      FC_W[1,9] := 0.25226828;
      FC_W[1,10] := -0.62714863;
      FC_W[1,11] := 0.07386149;
      FC_W[1,12] := -0.54759747;
      FC_W[1,13] := 0.00231634;
      FC_W[1,14] := -0.22999668;
      FC_W[1,15] := -0.03627737;
      FC_W[1,16] := -0.00447914;
      FC_W[1,17] := 0.00040707;
      FC_W[1,18] := 0.21295871;
      FC_W[1,19] := 0.21917404;
      FC_W[1,20] := -2.03310800;
      FC_W[1,21] := -0.23101221;
      FC_W[1,22] := 0.59129870;
      FC_W[1,23] := -0.14532049;
      FC_W[1,24] := 0.97670478;
      FC_W[1,25] := -0.18546271;
      FC_W[1,26] := 0.49225003;
      FC_W[1,27] := 0.23357685;
      FC_W[1,28] := -0.05720856;
      FC_W[1,29] := 0.13206857;
      FC_W[1,30] := 0.13029382;
      FC_W[1,31] := -0.28611091;
      FC_W[2,0] := -0.53158796;
      FC_W[2,1] := 2.18231130;
      FC_W[2,2] := 0.15426333;
      FC_W[2,3] := 0.93412578;
      FC_W[2,4] := 0.32678425;
      FC_W[2,5] := -0.29157385;
      FC_W[2,6] := -0.43484834;
      FC_W[2,7] := -0.40118921;
      FC_W[2,8] := -0.73715484;
      FC_W[2,9] := -1.47014546;
      FC_W[2,10] := 0.58461505;
      FC_W[2,11] := 0.72801095;
      FC_W[2,12] := -1.09524512;
      FC_W[2,13] := 0.17780326;
      FC_W[2,14] := 0.55109036;
      FC_W[2,15] := -0.46990421;
      FC_W[2,16] := -0.06730769;
      FC_W[2,17] := 0.69749105;
      FC_W[2,18] := 0.58266920;
      FC_W[2,19] := 0.02913308;
      FC_W[2,20] := 0.18312474;
      FC_W[2,21] := -0.12723203;
      FC_W[2,22] := 1.53492939;
      FC_W[2,23] := 1.18760669;
      FC_W[2,24] := -0.14219350;
      FC_W[2,25] := 0.37169734;
      FC_W[2,26] := -0.22027686;
      FC_W[2,27] := -0.33084327;
      FC_W[2,28] := -0.73663527;
      FC_W[2,29] := 0.07243921;
      FC_W[2,30] := 0.08782770;
      FC_W[2,31] := -0.84531319;
      FC_W[3,0] := 0.55170184;
      FC_W[3,1] := 2.12451887;
      FC_W[3,2] := -0.03638018;
      FC_W[3,3] := -0.92874491;
      FC_W[3,4] := 0.01098804;
      FC_W[3,5] := -0.12194143;
      FC_W[3,6] := -0.20283610;
      FC_W[3,7] := 0.71050656;
      FC_W[3,8] := -0.54710799;
      FC_W[3,9] := 0.84274971;
      FC_W[3,10] := -0.37954244;
      FC_W[3,11] := -0.17364120;
      FC_W[3,12] := 0.44716811;
      FC_W[3,13] := -0.05414552;
      FC_W[3,14] := -0.30617589;
      FC_W[3,15] := 0.00501720;
      FC_W[3,16] := -0.61364305;
      FC_W[3,17] := -0.40598497;
      FC_W[3,18] := 0.24112742;
      FC_W[3,19] := -0.18145135;
      FC_W[3,20] := 0.72023159;
      FC_W[3,21] := 0.31241485;
      FC_W[3,22] := -0.22940150;
      FC_W[3,23] := 0.32834825;
      FC_W[3,24] := -0.47077408;
      FC_W[3,25] := -0.41148546;
      FC_W[3,26] := 0.16142704;
      FC_W[3,27] := -0.05713443;
      FC_W[3,28] := -0.32514808;
      FC_W[3,29] := 0.26252571;
      FC_W[3,30] := 0.50961155;
      FC_W[3,31] := 0.53038257;
      FC_W[4,0] := -0.41400927;
      FC_W[4,1] := 1.33202946;
      FC_W[4,2] := 0.12711546;
      FC_W[4,3] := -0.08963529;
      FC_W[4,4] := 0.24866593;
      FC_W[4,5] := 0.08165067;
      FC_W[4,6] := 0.50525010;
      FC_W[4,7] := 0.82496148;
      FC_W[4,8] := 0.11588583;
      FC_W[4,9] := -0.21680501;
      FC_W[4,10] := 0.62970287;
      FC_W[4,11] := 0.06018925;
      FC_W[4,12] := 0.68656421;
      FC_W[4,13] := -1.21256888;
      FC_W[4,14] := -1.26492715;
      FC_W[4,15] := -0.70575857;
      FC_W[4,16] := -0.17878854;
      FC_W[4,17] := 0.27561840;
      FC_W[4,18] := -0.38193029;
      FC_W[4,19] := 0.25415263;
      FC_W[4,20] := -0.94903797;
      FC_W[4,21] := -0.59143215;
      FC_W[4,22] := -0.27362382;
      FC_W[4,23] := -0.23873141;
      FC_W[4,24] := -1.53285766;
      FC_W[4,25] := -0.27194324;
      FC_W[4,26] := -0.57270604;
      FC_W[4,27] := -0.31816959;
      FC_W[4,28] := 0.51076263;
      FC_W[4,29] := -0.39650953;
      FC_W[4,30] := -0.06086056;
      FC_W[4,31] := -0.04000641;
      FC_W[5,0] := 0.25593293;
      FC_W[5,1] := -0.71731991;
      FC_W[5,2] := 0.62669879;
      FC_W[5,3] := 1.38078809;
      FC_W[5,4] := -0.12516685;
      FC_W[5,5] := -0.90641493;
      FC_W[5,6] := -0.39019036;
      FC_W[5,7] := -0.45447922;
      FC_W[5,8] := 0.01198741;
      FC_W[5,9] := -0.21863569;
      FC_W[5,10] := 0.71772867;
      FC_W[5,11] := 0.27339056;
      FC_W[5,12] := 0.20110083;
      FC_W[5,13] := -0.13613328;
      FC_W[5,14] := -2.24843359;
      FC_W[5,15] := 0.12153642;
      FC_W[5,16] := 0.93278831;
      FC_W[5,17] := -0.95549434;
      FC_W[5,18] := 0.26438603;
      FC_W[5,19] := 0.19650064;
      FC_W[5,20] := -0.06620517;
      FC_W[5,21] := 0.29557747;
      FC_W[5,22] := 1.31400585;
      FC_W[5,23] := -0.15871854;
      FC_W[5,24] := 0.40522489;
      FC_W[5,25] := 0.03414011;
      FC_W[5,26] := -0.38867807;
      FC_W[5,27] := -0.81741858;
      FC_W[5,28] := 1.06798649;
      FC_W[5,29] := 3.75573659;
      FC_W[5,30] := -0.51656634;
      FC_W[5,31] := -0.28770104;
      FC_W[6,0] := -0.99143010;
      FC_W[6,1] := 0.29992977;
      FC_W[6,2] := 1.43284762;
      FC_W[6,3] := -0.34655777;
      FC_W[6,4] := -0.12928130;
      FC_W[6,5] := 0.15707546;
      FC_W[6,6] := -0.63261580;
      FC_W[6,7] := -0.29724568;
      FC_W[6,8] := 0.13134219;
      FC_W[6,9] := -1.04233253;
      FC_W[6,10] := 0.53604454;
      FC_W[6,11] := -0.18040322;
      FC_W[6,12] := 0.16615772;
      FC_W[6,13] := -0.40025923;
      FC_W[6,14] := -1.54933608;
      FC_W[6,15] := 0.41574958;
      FC_W[6,16] := 0.35386816;
      FC_W[6,17] := -0.45704508;
      FC_W[6,18] := 0.60151654;
      FC_W[6,19] := -0.67978704;
      FC_W[6,20] := 0.15072536;
      FC_W[6,21] := -0.42846721;
      FC_W[6,22] := -0.85208124;
      FC_W[6,23] := -0.05353868;
      FC_W[6,24] := 0.86764193;
      FC_W[6,25] := -0.24695079;
      FC_W[6,26] := 0.82921457;
      FC_W[6,27] := -1.08330154;
      FC_W[6,28] := 0.22054735;
      FC_W[6,29] := -0.23250555;
      FC_W[6,30] := 0.84133679;
      FC_W[6,31] := -0.10032179;
      FC_W[7,0] := 0.30265906;
      FC_W[7,1] := 2.08623362;
      FC_W[7,2] := 0.06350639;
      FC_W[7,3] := -1.09427238;
      FC_W[7,4] := -0.02930364;
      FC_W[7,5] := 0.24324393;
      FC_W[7,6] := 0.16107884;
      FC_W[7,7] := -0.00278581;
      FC_W[7,8] := 0.11302312;
      FC_W[7,9] := 0.10457820;
      FC_W[7,10] := -0.14860652;
      FC_W[7,11] := -0.10135441;
      FC_W[7,12] := 1.27947247;
      FC_W[7,13] := -0.08310315;
      FC_W[7,14] := -0.41487727;
      FC_W[7,15] := 0.17592667;
      FC_W[7,16] := -0.25739285;
      FC_W[7,17] := 0.24304490;
      FC_W[7,18] := -0.47447765;
      FC_W[7,19] := -0.28621474;
      FC_W[7,20] := 0.67906636;
      FC_W[7,21] := -0.40683922;
      FC_W[7,22] := -0.50886548;
      FC_W[7,23] := 0.06748977;
      FC_W[7,24] := -0.28961775;
      FC_W[7,25] := -0.11677405;
      FC_W[7,26] := 0.16660805;
      FC_W[7,27] := 0.34886500;
      FC_W[7,28] := -0.65834177;
      FC_W[7,29] := 0.30940986;
      FC_W[7,30] := -0.04497011;
      FC_W[7,31] := 0.22881326;
      FC_W[8,0] := 0.23515312;
      FC_W[8,1] := 2.35528612;
      FC_W[8,2] := 0.12001805;
      FC_W[8,3] := 0.60647392;
      FC_W[8,4] := -0.31542465;
      FC_W[8,5] := -0.26584071;
      FC_W[8,6] := 0.15293968;
      FC_W[8,7] := 0.19515641;
      FC_W[8,8] := -0.34400198;
      FC_W[8,9] := 0.12394456;
      FC_W[8,10] := 0.06283668;
      FC_W[8,11] := -0.67132694;
      FC_W[8,12] := -1.10496128;
      FC_W[8,13] := -0.33543864;
      FC_W[8,14] := 0.34250832;
      FC_W[8,15] := 0.11089487;
      FC_W[8,16] := 0.27817380;
      FC_W[8,17] := -0.27934778;
      FC_W[8,18] := 1.01753807;
      FC_W[8,19] := -0.14856282;
      FC_W[8,20] := 1.15498221;
      FC_W[8,21] := 0.31782010;
      FC_W[8,22] := -0.57135326;
      FC_W[8,23] := -0.27457404;
      FC_W[8,24] := -0.01912341;
      FC_W[8,25] := 0.07636409;
      FC_W[8,26] := -0.05262562;
      FC_W[8,27] := 0.01281669;
      FC_W[8,28] := 1.45306993;
      FC_W[8,29] := 0.01643326;
      FC_W[8,30] := 0.02226772;
      FC_W[8,31] := 0.16109315;
      FC_W[9,0] := 0.16771235;
      FC_W[9,1] := 2.17360902;
      FC_W[9,2] := 0.13744619;
      FC_W[9,3] := -0.45034087;
      FC_W[9,4] := -0.18103811;
      FC_W[9,5] := 0.19206211;
      FC_W[9,6] := 0.29432642;
      FC_W[9,7] := -0.29548097;
      FC_W[9,8] := 0.26934287;
      FC_W[9,9] := -0.23640421;
      FC_W[9,10] := 0.08889509;
      FC_W[9,11] := -0.29550803;
      FC_W[9,12] := 0.70984375;
      FC_W[9,13] := -0.18878627;
      FC_W[9,14] := -0.16082951;
      FC_W[9,15] := 0.28989646;
      FC_W[9,16] := 0.17481117;
      FC_W[9,17] := 0.31475934;
      FC_W[9,18] := -0.19749227;
      FC_W[9,19] := -0.29642978;
      FC_W[9,20] := 0.85720885;
      FC_W[9,21] := -0.43476731;
      FC_W[9,22] := -0.67719740;
      FC_W[9,23] := -0.20220257;
      FC_W[9,24] := -0.05126322;
      FC_W[9,25] := 0.10412872;
      FC_W[9,26] := 0.06379344;
      FC_W[9,27] := 0.43333077;
      FC_W[9,28] := 0.06093162;
      FC_W[9,29] := 0.21085459;
      FC_W[9,30] := -0.27212784;
      FC_W[9,31] := 0.04487327;
      FC_W[10,0] := 0.55635911;
      FC_W[10,1] := 1.71071684;
      FC_W[10,2] := -0.98758829;
      FC_W[10,3] := -1.20704234;
      FC_W[10,4] := 0.70373571;
      FC_W[10,5] := -0.49822235;
      FC_W[10,6] := -0.34963137;
      FC_W[10,7] := -0.04954350;
      FC_W[10,8] := 0.57998538;
      FC_W[10,9] := -0.12894104;
      FC_W[10,10] := 0.17007013;
      FC_W[10,11] := 0.22826548;
      FC_W[10,12] := 0.52343917;
      FC_W[10,13] := 0.24545214;
      FC_W[10,14] := 0.32942688;
      FC_W[10,15] := 0.31240448;
      FC_W[10,16] := -0.23860073;
      FC_W[10,17] := 0.84877467;
      FC_W[10,18] := -0.03334466;
      FC_W[10,19] := -0.08059564;
      FC_W[10,20] := -0.50759733;
      FC_W[10,21] := 0.57257271;
      FC_W[10,22] := -0.54642487;
      FC_W[10,23] := 0.07352713;
      FC_W[10,24] := 0.81966442;
      FC_W[10,25] := -0.40594006;
      FC_W[10,26] := -0.35969523;
      FC_W[10,27] := 1.14789081;
      FC_W[10,28] := 0.64354020;
      FC_W[10,29] := 1.38284671;
      FC_W[10,30] := -0.42893896;
      FC_W[10,31] := 0.09688565;
      FC_W[11,0] := -0.43645921;
      FC_W[11,1] := 0.23312488;
      FC_W[11,2] := -0.23381421;
      FC_W[11,3] := 1.35307658;
      FC_W[11,4] := 0.06825005;
      FC_W[11,5] := 0.04006363;
      FC_W[11,6] := -0.30487701;
      FC_W[11,7] := -0.04899468;
      FC_W[11,8] := -0.69408715;
      FC_W[11,9] := 0.32083067;
      FC_W[11,10] := -1.27051854;
      FC_W[11,11] := -0.28955328;
      FC_W[11,12] := 0.94128507;
      FC_W[11,13] := -0.04163137;
      FC_W[11,14] := -0.19035473;
      FC_W[11,15] := 1.00236845;
      FC_W[11,16] := 1.06163549;
      FC_W[11,17] := 0.45048153;
      FC_W[11,18] := 0.19175214;
      FC_W[11,19] := -0.00000184;
      FC_W[11,20] := -0.00385919;
      FC_W[11,21] := -0.25575012;
      FC_W[11,22] := 0.63028401;
      FC_W[11,23] := 0.23347531;
      FC_W[11,24] := 0.62187344;
      FC_W[11,25] := -0.06846938;
      FC_W[11,26] := -0.08085597;
      FC_W[11,27] := 0.08367075;
      FC_W[11,28] := 0.07401622;
      FC_W[11,29] := -0.68332726;
      FC_W[11,30] := 0.36182699;
      FC_W[11,31] := 0.09208941;
      FC_W[12,0] := -0.12697175;
      FC_W[12,1] := 0.54007989;
      FC_W[12,2] := -0.23235552;
      FC_W[12,3] := 1.02737308;
      FC_W[12,4] := -0.21164975;
      FC_W[12,5] := -0.18848586;
      FC_W[12,6] := -0.31116375;
      FC_W[12,7] := 0.18885162;
      FC_W[12,8] := 0.26512960;
      FC_W[12,9] := 0.64287508;
      FC_W[12,10] := 0.17899334;
      FC_W[12,11] := 0.11003251;
      FC_W[12,12] := 0.97311103;
      FC_W[12,13] := 0.04088512;
      FC_W[12,14] := 0.28795946;
      FC_W[12,15] := 1.57381439;
      FC_W[12,16] := 0.84596854;
      FC_W[12,17] := -0.53194338;
      FC_W[12,18] := 0.83031321;
      FC_W[12,19] := 0.19111450;
      FC_W[12,20] := -0.29391897;
      FC_W[12,21] := -0.53817254;
      FC_W[12,22] := 1.39124548;
      FC_W[12,23] := 0.21961257;
      FC_W[12,24] := 0.63080877;
      FC_W[12,25] := -0.13176970;
      FC_W[12,26] := 0.19578983;
      FC_W[12,27] := 0.07251017;
      FC_W[12,28] := 0.15489395;
      FC_W[12,29] := -0.56836164;
      FC_W[12,30] := 0.24469846;
      FC_W[12,31] := -0.29308897;
      FC_W[13,0] := 2.20791268;
      FC_W[13,1] := -1.10374355;
      FC_W[13,2] := -0.24162126;
      FC_W[13,3] := 0.77374041;
      FC_W[13,4] := -1.13711357;
      FC_W[13,5] := -1.31870210;
      FC_W[13,6] := 0.47841373;
      FC_W[13,7] := -0.16105147;
      FC_W[13,8] := -0.35249650;
      FC_W[13,9] := -0.42332867;
      FC_W[13,10] := -1.55202627;
      FC_W[13,11] := 1.01507616;
      FC_W[13,12] := -0.63866675;
      FC_W[13,13] := -0.71099406;
      FC_W[13,14] := -0.48592618;
      FC_W[13,15] := -0.37993100;
      FC_W[13,16] := 0.18940821;
      FC_W[13,17] := -0.05538184;
      FC_W[13,18] := -0.14446187;
      FC_W[13,19] := 0.44147074;
      FC_W[13,20] := -0.71370798;
      FC_W[13,21] := -1.35824025;
      FC_W[13,22] := -0.32107875;
      FC_W[13,23] := -0.66948777;
      FC_W[13,24] := 0.46409652;
      FC_W[13,25] := -0.56385392;
      FC_W[13,26] := 1.45479858;
      FC_W[13,27] := 1.22730565;
      FC_W[13,28] := -0.70979494;
      FC_W[13,29] := 0.23732866;
      FC_W[13,30] := 0.40240869;
      FC_W[13,31] := -0.91399556;
      FC_W[14,0] := -0.07104833;
      FC_W[14,1] := -0.28022146;
      FC_W[14,2] := -0.67785078;
      FC_W[14,3] := 0.19481595;
      FC_W[14,4] := -0.03060088;
      FC_W[14,5] := -0.20427652;
      FC_W[14,6] := 0.04726106;
      FC_W[14,7] := 1.98258340;
      FC_W[14,8] := 4.40404320;
      FC_W[14,9] := -1.24794614;
      FC_W[14,10] := -1.24316883;
      FC_W[14,11] := -1.68179226;
      FC_W[14,12] := -0.29661027;
      FC_W[14,13] := 0.01353078;
      FC_W[14,14] := -0.41424713;
      FC_W[14,15] := 0.58704215;
      FC_W[14,16] := -1.78230023;
      FC_W[14,17] := 1.53948402;
      FC_W[14,18] := -0.07893131;
      FC_W[14,19] := -3.22760653;
      FC_W[14,20] := 0.56132263;
      FC_W[14,21] := 0.12644786;
      FC_W[14,22] := 1.26095736;
      FC_W[14,23] := -0.00488345;
      FC_W[14,24] := 0.29457206;
      FC_W[14,25] := -1.28626144;
      FC_W[14,26] := -0.26738542;
      FC_W[14,27] := -0.44110236;
      FC_W[14,28] := -0.43122882;
      FC_W[14,29] := -0.00431219;
      FC_W[14,30] := -0.40952465;
      FC_W[14,31] := -0.30441639;
      FC_W[15,0] := 0.20250924;
      FC_W[15,1] := 0.43626478;
      FC_W[15,2] := 0.27463222;
      FC_W[15,3] := 0.37211508;
      FC_W[15,4] := -0.03340056;
      FC_W[15,5] := -0.06623933;
      FC_W[15,6] := -0.24864028;
      FC_W[15,7] := -0.58677751;
      FC_W[15,8] := -0.61499745;
      FC_W[15,9] := 0.54579276;
      FC_W[15,10] := -0.19726747;
      FC_W[15,11] := 0.12831730;
      FC_W[15,12] := 0.61062902;
      FC_W[15,13] := -0.02127237;
      FC_W[15,14] := 0.21842071;
      FC_W[15,15] := -0.17562330;
      FC_W[15,16] := 0.38656747;
      FC_W[15,17] := 0.59372723;
      FC_W[15,18] := 0.24492693;
      FC_W[15,19] := -1.01225615;
      FC_W[15,20] := -0.01717149;
      FC_W[15,21] := 0.54135400;
      FC_W[15,22] := 1.04819000;
      FC_W[15,23] := -1.09988487;
      FC_W[15,24] := -0.29471993;
      FC_W[15,25] := 0.78609461;
      FC_W[15,26] := 0.23125337;
      FC_W[15,27] := -0.02700599;
      FC_W[15,28] := 0.42768958;
      FC_W[15,29] := -0.29631129;
      FC_W[15,30] := 1.83250082;
      FC_W[15,31] := -0.43059009;
      FC_W[16,0] := -0.37697601;
      FC_W[16,1] := -0.19721903;
      FC_W[16,2] := -0.13793600;
      FC_W[16,3] := 0.07084525;
      FC_W[16,4] := 0.47389659;
      FC_W[16,5] := 0.68528003;
      FC_W[16,6] := 1.65266597;
      FC_W[16,7] := -0.24744993;
      FC_W[16,8] := 1.25457382;
      FC_W[16,9] := 1.49639773;
      FC_W[16,10] := 0.50168604;
      FC_W[16,11] := -0.50251526;
      FC_W[16,12] := -0.00292949;
      FC_W[16,13] := -0.70094889;
      FC_W[16,14] := 0.17360571;
      FC_W[16,15] := -0.58291054;
      FC_W[16,16] := 0.50401050;
      FC_W[16,17] := -1.54409647;
      FC_W[16,18] := -1.89241540;
      FC_W[16,19] := -0.33420387;
      FC_W[16,20] := 0.63442737;
      FC_W[16,21] := -0.10250572;
      FC_W[16,22] := -0.74442780;
      FC_W[16,23] := 2.23745084;
      FC_W[16,24] := 0.97562188;
      FC_W[16,25] := -0.53874046;
      FC_W[16,26] := 0.44360429;
      FC_W[16,27] := 0.48179910;
      FC_W[16,28] := 1.56847930;
      FC_W[16,29] := 0.12322044;
      FC_W[16,30] := 0.58041352;
      FC_W[16,31] := -2.92400813;
      FC_W[17,0] := -0.28855094;
      FC_W[17,1] := -0.73520070;
      FC_W[17,2] := -0.58204508;
      FC_W[17,3] := -2.53923368;
      FC_W[17,4] := 0.04207829;
      FC_W[17,5] := 0.34026721;
      FC_W[17,6] := 0.83833164;
      FC_W[17,7] := 1.37610734;
      FC_W[17,8] := -0.48114690;
      FC_W[17,9] := 0.80318284;
      FC_W[17,10] := 1.40226424;
      FC_W[17,11] := 1.19034028;
      FC_W[17,12] := -1.82810128;
      FC_W[17,13] := 0.07092776;
      FC_W[17,14] := -0.24957196;
      FC_W[17,15] := 0.41651461;
      FC_W[17,16] := 2.31544805;
      FC_W[17,17] := -0.29625085;
      FC_W[17,18] := 0.43194380;
      FC_W[17,19] := -2.91967225;
      FC_W[17,20] := 0.48595843;
      FC_W[17,21] := -0.95144910;
      FC_W[17,22] := -0.56275243;
      FC_W[17,23] := 0.17238346;
      FC_W[17,24] := 0.18526348;
      FC_W[17,25] := -1.61428738;
      FC_W[17,26] := -0.85377961;
      FC_W[17,27] := -0.13946605;
      FC_W[17,28] := -0.68767577;
      FC_W[17,29] := 0.88757920;
      FC_W[17,30] := -1.37992692;
      FC_W[17,31] := -0.30283210;
      FC_W[18,0] := -0.60211664;
      FC_W[18,1] := -0.47432238;
      FC_W[18,2] := 0.49715492;
      FC_W[18,3] := -1.05803704;
      FC_W[18,4] := 0.31516069;
      FC_W[18,5] := 0.60292727;
      FC_W[18,6] := -1.12411284;
      FC_W[18,7] := -0.81225699;
      FC_W[18,8] := 0.22442850;
      FC_W[18,9] := -0.31069636;
      FC_W[18,10] := -0.39883116;
      FC_W[18,11] := -0.00383187;
      FC_W[18,12] := -1.32017577;
      FC_W[18,13] := 0.76117158;
      FC_W[18,14] := -0.59863925;
      FC_W[18,15] := 2.91382790;
      FC_W[18,16] := -0.31635019;
      FC_W[18,17] := -0.69926184;
      FC_W[18,18] := 0.44085792;
      FC_W[18,19] := -0.27446097;
      FC_W[18,20] := 0.68643546;
      FC_W[18,21] := -1.84294975;
      FC_W[18,22] := -0.20962636;
      FC_W[18,23] := -0.22959881;
      FC_W[18,24] := 0.18067747;
      FC_W[18,25] := 0.47698760;
      FC_W[18,26] := -3.78073096;
      FC_W[18,27] := 0.82570255;
      FC_W[18,28] := -0.23815499;
      FC_W[18,29] := 1.09470105;
      FC_W[18,30] := 1.66854107;
      FC_W[18,31] := -0.13462155;
      FC_W[19,0] := 0.44800782;
      FC_W[19,1] := 0.06498748;
      FC_W[19,2] := -0.06952048;
      FC_W[19,3] := -0.51742721;
      FC_W[19,4] := -0.09736256;
      FC_W[19,5] := -0.37422362;
      FC_W[19,6] := -0.15245904;
      FC_W[19,7] := 0.63320434;
      FC_W[19,8] := 1.04222059;
      FC_W[19,9] := 0.06480665;
      FC_W[19,10] := 0.35045585;
      FC_W[19,11] := -0.40922517;
      FC_W[19,12] := -0.08025740;
      FC_W[19,13] := 0.05562712;
      FC_W[19,14] := 0.10890836;
      FC_W[19,15] := -0.13707444;
      FC_W[19,16] := 1.62350214;
      FC_W[19,17] := 0.41023293;
      FC_W[19,18] := 0.34094810;
      FC_W[19,19] := 0.31232962;
      FC_W[19,20] := -0.14682344;
      FC_W[19,21] := 0.48118156;
      FC_W[19,22] := 0.78214991;
      FC_W[19,23] := 0.03551027;
      FC_W[19,24] := -0.44571006;
      FC_W[19,25] := -0.08649512;
      FC_W[19,26] := 0.47158131;
      FC_W[19,27] := -0.36406398;
      FC_W[19,28] := -0.22915788;
      FC_W[19,29] := 0.01263516;
      FC_W[19,30] := 0.57616603;
      FC_W[19,31] := 0.12845607;
      FC_W[20,0] := 0.55101711;
      FC_W[20,1] := 0.35684553;
      FC_W[20,2] := -0.92210096;
      FC_W[20,3] := 0.13750382;
      FC_W[20,4] := 0.01511240;
      FC_W[20,5] := -0.63257527;
      FC_W[20,6] := 1.40384579;
      FC_W[20,7] := -0.21248135;
      FC_W[20,8] := -0.16805060;
      FC_W[20,9] := -0.11867571;
      FC_W[20,10] := -0.39359516;
      FC_W[20,11] := -0.15843204;
      FC_W[20,12] := 0.22070603;
      FC_W[20,13] := 0.71381277;
      FC_W[20,14] := -0.11454471;
      FC_W[20,15] := -0.38763249;
      FC_W[20,16] := -0.09213293;
      FC_W[20,17] := -0.03829917;
      FC_W[20,18] := -0.25112540;
      FC_W[20,19] := 0.09202781;
      FC_W[20,20] := -0.79897386;
      FC_W[20,21] := 0.14058812;
      FC_W[20,22] := -0.30311379;
      FC_W[20,23] := -0.43297794;
      FC_W[20,24] := 0.11171950;
      FC_W[20,25] := 0.17598327;
      FC_W[20,26] := -0.82704544;
      FC_W[20,27] := -0.20293660;
      FC_W[20,28] := -0.50960398;
      FC_W[20,29] := -0.13715295;
      FC_W[20,30] := -0.20570764;
      FC_W[20,31] := -0.22419536;
      FC_W[21,0] := -1.38703454;
      FC_W[21,1] := 0.13443221;
      FC_W[21,2] := 1.65575707;
      FC_W[21,3] := -0.30523026;
      FC_W[21,4] := 0.20814605;
      FC_W[21,5] := 0.44282535;
      FC_W[21,6] := -0.18247518;
      FC_W[21,7] := 0.68251020;
      FC_W[21,8] := -0.51809436;
      FC_W[21,9] := -0.59682101;
      FC_W[21,10] := 0.32860571;
      FC_W[21,11] := -0.65614474;
      FC_W[21,12] := -0.12320014;
      FC_W[21,13] := 1.67703843;
      FC_W[21,14] := 0.01895689;
      FC_W[21,15] := 0.41568109;
      FC_W[21,16] := 0.12311991;
      FC_W[21,17] := -0.85774213;
      FC_W[21,18] := -0.30047303;
      FC_W[21,19] := -0.33377433;
      FC_W[21,20] := 0.02386909;
      FC_W[21,21] := -0.03189978;
      FC_W[21,22] := 0.33781007;
      FC_W[21,23] := -0.20913075;
      FC_W[21,24] := -0.16453424;
      FC_W[21,25] := -0.14679955;
      FC_W[21,26] := 0.59973520;
      FC_W[21,27] := 0.48085397;
      FC_W[21,28] := 0.24753553;
      FC_W[21,29] := -0.01857807;
      FC_W[21,30] := 0.12446254;
      FC_W[21,31] := 0.10629370;
      FC_W[22,0] := 0.19716617;
      FC_W[22,1] := 0.13620606;
      FC_W[22,2] := 0.04876109;
      FC_W[22,3] := 0.23500557;
      FC_W[22,4] := 0.64577067;
      FC_W[22,5] := 0.25040030;
      FC_W[22,6] := 0.29043925;
      FC_W[22,7] := 0.85402560;
      FC_W[22,8] := 0.06459093;
      FC_W[22,9] := -1.23667681;
      FC_W[22,10] := -0.05787567;
      FC_W[22,11] := 0.74056232;
      FC_W[22,12] := 0.22630619;
      FC_W[22,13] := -0.10364483;
      FC_W[22,14] := -0.08892694;
      FC_W[22,15] := -0.34050211;
      FC_W[22,16] := 0.65094274;
      FC_W[22,17] := -1.17275202;
      FC_W[22,18] := -0.78813517;
      FC_W[22,19] := 0.34167442;
      FC_W[22,20] := 0.37342751;
      FC_W[22,21] := 0.12655480;
      FC_W[22,22] := 0.14093940;
      FC_W[22,23] := -0.97658986;
      FC_W[22,24] := 0.29666159;
      FC_W[22,25] := -0.95207864;
      FC_W[22,26] := -0.25645512;
      FC_W[22,27] := 0.21099935;
      FC_W[22,28] := -0.17070027;
      FC_W[22,29] := -0.15547353;
      FC_W[22,30] := 0.05844394;
      FC_W[22,31] := -0.35387653;
      FC_W[23,0] := 2.36117458;
      FC_W[23,1] := -0.27253562;
      FC_W[23,2] := -0.44734445;
      FC_W[23,3] := 0.43230754;
      FC_W[23,4] := 2.77088666;
      FC_W[23,5] := -1.15746760;
      FC_W[23,6] := -0.15780434;
      FC_W[23,7] := -0.08052579;
      FC_W[23,8] := -1.13770092;
      FC_W[23,9] := 0.34222582;
      FC_W[23,10] := -0.76248449;
      FC_W[23,11] := -0.31606591;
      FC_W[23,12] := -0.26905468;
      FC_W[23,13] := -0.65461212;
      FC_W[23,14] := 0.29336941;
      FC_W[23,15] := -0.56090289;
      FC_W[23,16] := -0.30688983;
      FC_W[23,17] := 0.29983157;
      FC_W[23,18] := -0.73118234;
      FC_W[23,19] := -0.10799882;
      FC_W[23,20] := -0.22133076;
      FC_W[23,21] := -1.62908876;
      FC_W[23,22] := 0.32420984;
      FC_W[23,23] := 0.12469828;
      FC_W[23,24] := 0.86695164;
      FC_W[23,25] := 0.00903137;
      FC_W[23,26] := 1.11415207;
      FC_W[23,27] := -0.62709349;
      FC_W[23,28] := -0.02971547;
      FC_W[23,29] := -0.25179407;
      FC_W[23,30] := -0.06880520;
      FC_W[23,31] := 0.58122498;
      FC_W[24,0] := 0.07595386;
      FC_W[24,1] := 0.17389667;
      FC_W[24,2] := -0.13460560;
      FC_W[24,3] := 0.23620439;
      FC_W[24,4] := 0.71178508;
      FC_W[24,5] := 0.42975000;
      FC_W[24,6] := 0.46598688;
      FC_W[24,7] := 1.36021495;
      FC_W[24,8] := 0.10479560;
      FC_W[24,9] := -0.78181171;
      FC_W[24,10] := -0.17630832;
      FC_W[24,11] := 0.88054228;
      FC_W[24,12] := 0.23260193;
      FC_W[24,13] := -0.07906808;
      FC_W[24,14] := 0.03967582;
      FC_W[24,15] := -0.41637811;
      FC_W[24,16] := 0.38345000;
      FC_W[24,17] := -0.55840528;
      FC_W[24,18] := -0.90066504;
      FC_W[24,19] := 0.97068053;
      FC_W[24,20] := 0.60454738;
      FC_W[24,21] := 0.02299176;
      FC_W[24,22] := 0.09866967;
      FC_W[24,23] := -1.46094978;
      FC_W[24,24] := 0.38187879;
      FC_W[24,25] := -1.42997479;
      FC_W[24,26] := -0.37488067;
      FC_W[24,27] := -0.04411485;
      FC_W[24,28] := -0.29138446;
      FC_W[24,29] := -0.07532097;
      FC_W[24,30] := -0.00954079;
      FC_W[24,31] := -0.99948364;
      FC_W[25,0] := 0.08445936;
      FC_W[25,1] := 0.16368021;
      FC_W[25,2] := -0.11429817;
      FC_W[25,3] := 0.25485840;
      FC_W[25,4] := 0.72819227;
      FC_W[25,5] := 0.42307603;
      FC_W[25,6] := 0.45525894;
      FC_W[25,7] := 1.32385421;
      FC_W[25,8] := 0.11924174;
      FC_W[25,9] := -0.79466659;
      FC_W[25,10] := -0.16143492;
      FC_W[25,11] := 0.87378216;
      FC_W[25,12] := 0.22462815;
      FC_W[25,13] := -0.08033443;
      FC_W[25,14] := 0.01655862;
      FC_W[25,15] := -0.40789300;
      FC_W[25,16] := 0.40738490;
      FC_W[25,17] := -0.57628548;
      FC_W[25,18] := -0.88914770;
      FC_W[25,19] := 0.94886303;
      FC_W[25,20] := 0.60112166;
      FC_W[25,21] := 0.02799439;
      FC_W[25,22] := 0.08625803;
      FC_W[25,23] := -1.44966817;
      FC_W[25,24] := 0.37795368;
      FC_W[25,25] := -1.41334343;
      FC_W[25,26] := -0.38357916;
      FC_W[25,27] := -0.01546234;
      FC_W[25,28] := -0.29737470;
      FC_W[25,29] := -0.08744591;
      FC_W[25,30] := -0.01248721;
      FC_W[25,31] := -0.99227226;
      FC_W[26,0] := 2.38675141;
      FC_W[26,1] := 0.10531798;
      FC_W[26,2] := 0.00214429;
      FC_W[26,3] := 0.29302251;
      FC_W[26,4] := -0.95878249;
      FC_W[26,5] := -0.62310410;
      FC_W[26,6] := -0.31759438;
      FC_W[26,7] := 0.11338235;
      FC_W[26,8] := -0.31615138;
      FC_W[26,9] := -1.49054682;
      FC_W[26,10] := 0.93792856;
      FC_W[26,11] := 0.87154341;
      FC_W[26,12] := 0.41643369;
      FC_W[26,13] := -1.12895298;
      FC_W[26,14] := -0.42944503;
      FC_W[26,15] := -0.59216714;
      FC_W[26,16] := 0.45720932;
      FC_W[26,17] := -0.10903971;
      FC_W[26,18] := -1.34624648;
      FC_W[26,19] := -0.30879995;
      FC_W[26,20] := 0.24794732;
      FC_W[26,21] := 0.29367086;
      FC_W[26,22] := 0.73384720;
      FC_W[26,23] := 0.23941633;
      FC_W[26,24] := 0.97845572;
      FC_W[26,25] := -0.83140624;
      FC_W[26,26] := -1.05813015;
      FC_W[26,27] := -0.12844378;
      FC_W[26,28] := 0.53951097;
      FC_W[26,29] := -0.46631601;
      FC_W[26,30] := -0.12978332;
      FC_W[26,31] := 0.57293302;
      FC_W[27,0] := -0.82125789;
      FC_W[27,1] := 0.24535166;
      FC_W[27,2] := 2.14815331;
      FC_W[27,3] := 0.07394390;
      FC_W[27,4] := 0.37535343;
      FC_W[27,5] := 0.20946552;
      FC_W[27,6] := -0.22952469;
      FC_W[27,7] := 0.21198778;
      FC_W[27,8] := 0.45519185;
      FC_W[27,9] := 0.43655413;
      FC_W[27,10] := 0.14163223;
      FC_W[27,11] := 0.37753379;
      FC_W[27,12] := -0.03609978;
      FC_W[27,13] := 1.92808294;
      FC_W[27,14] := 0.01438947;
      FC_W[27,15] := 0.12405793;
      FC_W[27,16] := 0.13592151;
      FC_W[27,17] := 0.25425518;
      FC_W[27,18] := -0.02739565;
      FC_W[27,19] := -0.02477069;
      FC_W[27,20] := 0.06481469;
      FC_W[27,21] := 0.01653567;
      FC_W[27,22] := -0.02758124;
      FC_W[27,23] := 0.17188995;
      FC_W[27,24] := -0.64550167;
      FC_W[27,25] := -0.43979689;
      FC_W[27,26] := 0.12660854;
      FC_W[27,27] := 0.10706360;
      FC_W[27,28] := 0.51992017;
      FC_W[27,29] := -0.04491308;
      FC_W[27,30] := 0.01514542;
      FC_W[27,31] := 0.33560848;
      FC_W[28,0] := -0.04899776;
      FC_W[28,1] := 0.30701822;
      FC_W[28,2] := 1.92029631;
      FC_W[28,3] := 0.04663092;
      FC_W[28,4] := 0.13275446;
      FC_W[28,5] := -0.48249826;
      FC_W[28,6] := 0.35161558;
      FC_W[28,7] := 0.07966720;
      FC_W[28,8] := -0.07919965;
      FC_W[28,9] := 0.38876459;
      FC_W[28,10] := -0.17509958;
      FC_W[28,11] := -0.39602360;
      FC_W[28,12] := 0.15088342;
      FC_W[28,13] := -1.95759904;
      FC_W[28,14] := 0.18524067;
      FC_W[28,15] := -0.07970117;
      FC_W[28,16] := 0.11674451;
      FC_W[28,17] := -0.51323682;
      FC_W[28,18] := 0.00075771;
      FC_W[28,19] := -0.21001135;
      FC_W[28,20] := -0.75531536;
      FC_W[28,21] := -0.03187747;
      FC_W[28,22] := 0.17554842;
      FC_W[28,23] := -0.06124675;
      FC_W[28,24] := -0.49238649;
      FC_W[28,25] := -0.42485896;
      FC_W[28,26] := -0.15337357;
      FC_W[28,27] := 0.14139321;
      FC_W[28,28] := -0.23361476;
      FC_W[28,29] := -0.02120185;
      FC_W[28,30] := -0.10555608;
      FC_W[28,31] := 0.25831261;
      FC_W[29,0] := 0.17467082;
      FC_W[29,1] := -1.15403891;
      FC_W[29,2] := 0.42410749;
      FC_W[29,3] := 0.68594784;
      FC_W[29,4] := 1.10142064;
      FC_W[29,5] := -0.02245768;
      FC_W[29,6] := 0.48027182;
      FC_W[29,7] := -0.64551872;
      FC_W[29,8] := -0.18186948;
      FC_W[29,9] := 1.84850705;
      FC_W[29,10] := 2.83370781;
      FC_W[29,11] := -1.14294016;
      FC_W[29,12] := -0.72066194;
      FC_W[29,13] := -0.59360534;
      FC_W[29,14] := -3.17248583;
      FC_W[29,15] := 0.69748610;
      FC_W[29,16] := -1.15201128;
      FC_W[29,17] := 1.43731534;
      FC_W[29,18] := 0.86861062;
      FC_W[29,19] := 0.54476595;
      FC_W[29,20] := 0.31251097;
      FC_W[29,21] := 0.58345324;
      FC_W[29,22] := 0.32586187;
      FC_W[29,23] := -0.83482420;
      FC_W[29,24] := 0.36158529;
      FC_W[29,25] := -0.74989313;
      FC_W[29,26] := 0.24822375;
      FC_W[29,27] := 2.35983777;
      FC_W[29,28] := -1.56794560;
      FC_W[29,29] := -1.44592392;
      FC_W[29,30] := -0.02158822;
      FC_W[29,31] := -1.23422480;
      FC_W[30,0] := 0.19600290;
      FC_W[30,1] := 0.13682650;
      FC_W[30,2] := 0.04799474;
      FC_W[30,3] := 0.23437470;
      FC_W[30,4] := 0.64216888;
      FC_W[30,5] := 0.24906796;
      FC_W[30,6] := 0.29510096;
      FC_W[30,7] := 0.85068154;
      FC_W[30,8] := 0.06323259;
      FC_W[30,9] := -1.24682426;
      FC_W[30,10] := -0.05564035;
      FC_W[30,11] := 0.73768073;
      FC_W[30,12] := 0.22608444;
      FC_W[30,13] := -0.10548198;
      FC_W[30,14] := -0.08953846;
      FC_W[30,15] := -0.34236404;
      FC_W[30,16] := 0.65254492;
      FC_W[30,17] := -1.17795432;
      FC_W[30,18] := -0.79025835;
      FC_W[30,19] := 0.33610207;
      FC_W[30,20] := 0.37127289;
      FC_W[30,21] := 0.12772927;
      FC_W[30,22] := 0.14501528;
      FC_W[30,23] := -0.96899563;
      FC_W[30,24] := 0.29870170;
      FC_W[30,25] := -0.94649816;
      FC_W[30,26] := -0.25102472;
      FC_W[30,27] := 0.21240576;
      FC_W[30,28] := -0.16554664;
      FC_W[30,29] := -0.15445521;
      FC_W[30,30] := 0.05736541;
      FC_W[30,31] := -0.34062430;
      FC_W[31,0] := -0.06291415;
      FC_W[31,1] := -0.13268666;
      FC_W[31,2] := 0.14153177;
      FC_W[31,3] := 0.05869582;
      FC_W[31,4] := 0.98602140;
      FC_W[31,5] := 0.33257216;
      FC_W[31,6] := 1.13677454;
      FC_W[31,7] := 0.49982995;
      FC_W[31,8] := 0.51303792;
      FC_W[31,9] := -1.36589992;
      FC_W[31,10] := -0.18576875;
      FC_W[31,11] := 1.36524236;
      FC_W[31,12] := -0.04106874;
      FC_W[31,13] := -0.35705602;
      FC_W[31,14] := -0.11357384;
      FC_W[31,15] := -0.45420462;
      FC_W[31,16] := 0.65129673;
      FC_W[31,17] := -1.11419582;
      FC_W[31,18] := -0.32770509;
      FC_W[31,19] := 0.44034311;
      FC_W[31,20] := 0.59986246;
      FC_W[31,21] := 0.21020119;
      FC_W[31,22] := 0.25237066;
      FC_W[31,23] := -0.75997669;
      FC_W[31,24] := 0.35624456;
      FC_W[31,25] := -0.91603827;
      FC_W[31,26] := 0.02340161;
      FC_W[31,27] := 0.28168905;
      FC_W[31,28] := 0.09072609;
      FC_W[31,29] := 0.00274630;
      FC_W[31,30] := 0.38698420;
      FC_W[31,31] := 0.65330857;
      FC_W[32,0] := 0.45316526;
      FC_W[32,1] := 0.21850894;
      FC_W[32,2] := 0.43266058;
      FC_W[32,3] := 0.53624105;
      FC_W[32,4] := 0.78354108;
      FC_W[32,5] := 0.07270878;
      FC_W[32,6] := -0.41047511;
      FC_W[32,7] := 0.34728459;
      FC_W[32,8] := 0.42241964;
      FC_W[32,9] := -1.07310939;
      FC_W[32,10] := -0.29135448;
      FC_W[32,11] := 0.73983669;
      FC_W[32,12] := 0.36980560;
      FC_W[32,13] := 0.16045348;
      FC_W[32,14] := -0.16240825;
      FC_W[32,15] := -0.27712277;
      FC_W[32,16] := 1.10141444;
      FC_W[32,17] := -1.58855307;
      FC_W[32,18] := -0.63992548;
      FC_W[32,19] := -0.16592859;
      FC_W[32,20] := 0.04723974;
      FC_W[32,21] := 0.22148028;
      FC_W[32,22] := -0.32578921;
      FC_W[32,23] := -0.57134801;
      FC_W[32,24] := -0.10733084;
      FC_W[32,25] := -0.54068953;
      FC_W[32,26] := -0.41983676;
      FC_W[32,27] := 0.24719903;
      FC_W[32,28] := -0.28076965;
      FC_W[32,29] := -0.25654367;
      FC_W[32,30] := -0.05608768;
      FC_W[32,31] := -0.33111042;
      FC_W[33,0] := 0.58171481;
      FC_W[33,1] := 0.28558809;
      FC_W[33,2] := 0.70109051;
      FC_W[33,3] := 0.52311713;
      FC_W[33,4] := 0.56277329;
      FC_W[33,5] := -0.12312344;
      FC_W[33,6] := -0.81610090;
      FC_W[33,7] := -0.19942789;
      FC_W[33,8] := 0.48381969;
      FC_W[33,9] := -1.49506116;
      FC_W[33,10] := -0.36867550;
      FC_W[33,11] := 0.64773238;
      FC_W[33,12] := 0.46802661;
      FC_W[33,13] := 0.25560713;
      FC_W[33,14] := -0.13315524;
      FC_W[33,15] := -0.22961804;
      FC_W[33,16] := 1.48115480;
      FC_W[33,17] := -2.24376726;
      FC_W[33,18] := -0.54044688;
      FC_W[33,19] := -0.91481858;
      FC_W[33,20] := -0.28749046;
      FC_W[33,21] := 0.36017141;
      FC_W[33,22] := -0.43211988;
      FC_W[33,23] := 0.09178846;
      FC_W[33,24] := -0.34466580;
      FC_W[33,25] := 0.06815648;
      FC_W[33,26] := -0.37362421;
      FC_W[33,27] := 0.32526520;
      FC_W[33,28] := -0.09456850;
      FC_W[33,29] := -0.27243760;
      FC_W[33,30] := -0.02762402;
      FC_W[33,31] := 0.35988516;
      FC_W[34,0] := 0.39796761;
      FC_W[34,1] := 0.34505269;
      FC_W[34,2] := 0.42251158;
      FC_W[34,3] := 0.37203887;
      FC_W[34,4] := 0.42278188;
      FC_W[34,5] := -0.03246171;
      FC_W[34,6] := -0.55399013;
      FC_W[34,7] := 0.12313119;
      FC_W[34,8] := 0.27692446;
      FC_W[34,9] := -1.58456337;
      FC_W[34,10] := -0.35354123;
      FC_W[34,11] := 0.61738098;
      FC_W[34,12] := 0.42633978;
      FC_W[34,13] := 0.18016912;
      FC_W[34,14] := 0.03770608;
      FC_W[34,15] := -0.26501924;
      FC_W[34,16] := 1.24879241;
      FC_W[34,17] := -2.01006579;
      FC_W[34,18] := -0.61255771;
      FC_W[34,19] := -0.64846724;
      FC_W[34,20] := -0.15543117;
      FC_W[34,21] := 0.23150840;
      FC_W[34,22] := -0.25104845;
      FC_W[34,23] := -0.13263990;
      FC_W[34,24] := -0.17177737;
      FC_W[34,25] := -0.08472409;
      FC_W[34,26] := -0.30952516;
      FC_W[34,27] := 0.14638457;
      FC_W[34,28] := 0.01033866;
      FC_W[34,29] := -0.17122130;
      FC_W[34,30] := 0.00483797;
      FC_W[34,31] := 0.21764055;
      FC_W[35,0] := 0.47281465;
      FC_W[35,1] := 0.22640406;
      FC_W[35,2] := 0.37663290;
      FC_W[35,3] := 0.64435512;
      FC_W[35,4] := 0.99040037;
      FC_W[35,5] := 0.11951960;
      FC_W[35,6] := -0.41641048;
      FC_W[35,7] := 0.55413467;
      FC_W[35,8] := 0.46428216;
      FC_W[35,9] := -0.70929921;
      FC_W[35,10] := -0.36132902;
      FC_W[35,11] := 0.75798023;
      FC_W[35,12] := 0.35432577;
      FC_W[35,13] := 0.20557950;
      FC_W[35,14] := -0.18643822;
      FC_W[35,15] := -0.29398799;
      FC_W[35,16] := 0.99243772;
      FC_W[35,17] := -1.27834427;
      FC_W[35,18] := -0.66676456;
      FC_W[35,19] := 0.13668784;
      FC_W[35,20] := 0.11368812;
      FC_W[35,21] := 0.11678398;
      FC_W[35,22] := -0.43666810;
      FC_W[35,23] := -0.84696633;
      FC_W[35,24] := -0.09376711;
      FC_W[35,25] := -0.74521321;
      FC_W[35,26] := -0.47813976;
      FC_W[35,27] := 0.15896457;
      FC_W[35,28] := -0.41975939;
      FC_W[35,29] := -0.27025852;
      FC_W[35,30] := -0.12737930;
      FC_W[35,31] := -0.78730679;
      FC_W[36,0] := -0.27766651;
      FC_W[36,1] := -0.11740696;
      FC_W[36,2] := -1.31230485;
      FC_W[36,3] := 0.12661482;
      FC_W[36,4] := 0.02779600;
      FC_W[36,5] := 0.53574544;
      FC_W[36,6] := 0.10322278;
      FC_W[36,7] := -1.33259964;
      FC_W[36,8] := -0.16246226;
      FC_W[36,9] := -0.76596600;
      FC_W[36,10] := -0.07376932;
      FC_W[36,11] := -0.38214219;
      FC_W[36,12] := -0.00662602;
      FC_W[36,13] := 0.90929550;
      FC_W[36,14] := -0.01971030;
      FC_W[36,15] := -0.40236777;
      FC_W[36,16] := 0.24568664;
      FC_W[36,17] := -0.45955896;
      FC_W[36,18] := -0.12628753;
      FC_W[36,19] := 0.45840219;
      FC_W[36,20] := 0.28605455;
      FC_W[36,21] := -0.28069675;
      FC_W[36,22] := 0.05465906;
      FC_W[36,23] := -0.95575094;
      FC_W[36,24] := -1.59583950;
      FC_W[36,25] := -3.89907908;
      FC_W[36,26] := 0.13362858;
      FC_W[36,27] := 0.00279548;
      FC_W[36,28] := -0.36037770;
      FC_W[36,29] := -0.02456625;
      FC_W[36,30] := 0.03994703;
      FC_W[36,31] := -0.84338814;
      FC_W[37,0] := 0.48596013;
      FC_W[37,1] := 0.21791193;
      FC_W[37,2] := 0.37341836;
      FC_W[37,3] := 0.67805314;
      FC_W[37,4] := 1.04353714;
      FC_W[37,5] := 0.13452934;
      FC_W[37,6] := -0.41462234;
      FC_W[37,7] := 0.59311748;
      FC_W[37,8] := 0.48404527;
      FC_W[37,9] := -0.61081266;
      FC_W[37,10] := -0.37112591;
      FC_W[37,11] := 0.77415752;
      FC_W[37,12] := 0.34494308;
      FC_W[37,13] := 0.21793722;
      FC_W[37,14] := -0.19704254;
      FC_W[37,15] := -0.29635364;
      FC_W[37,16] := 0.96507460;
      FC_W[37,17] := -1.18958211;
      FC_W[37,18] := -0.66671556;
      FC_W[37,19] := 0.21892339;
      FC_W[37,20] := 0.13998653;
      FC_W[37,21] := 0.09513262;
      FC_W[37,22] := -0.45922533;
      FC_W[37,23] := -0.91865146;
      FC_W[37,24] := -0.08645191;
      FC_W[37,25] := -0.82173491;
      FC_W[37,26] := -0.48824522;
      FC_W[37,27] := 0.14734998;
      FC_W[37,28] := -0.45822144;
      FC_W[37,29] := -0.27875769;
      FC_W[37,30] := -0.14206089;
      FC_W[37,31] := -0.90061128;
      FC_W[38,0] := 0.90194970;
      FC_W[38,1] := -0.02848357;
      FC_W[38,2] := 0.24474472;
      FC_W[38,3] := -0.77616340;
      FC_W[38,4] := 0.38411501;
      FC_W[38,5] := -0.13671793;
      FC_W[38,6] := 1.00297904;
      FC_W[38,7] := 0.34290555;
      FC_W[38,8] := -0.66706288;
      FC_W[38,9] := -0.96812254;
      FC_W[38,10] := 0.51059961;
      FC_W[38,11] := 0.30854204;
      FC_W[38,12] := -0.35195786;
      FC_W[38,13] := -0.37104955;
      FC_W[38,14] := 0.26861626;
      FC_W[38,15] := 3.64562392;
      FC_W[38,16] := -0.76310056;
      FC_W[38,17] := 0.33728310;
      FC_W[38,18] := -1.09334779;
      FC_W[38,19] := -0.57048130;
      FC_W[38,20] := 0.07434628;
      FC_W[38,21] := 1.44640696;
      FC_W[38,22] := -0.69001889;
      FC_W[38,23] := 0.59528297;
      FC_W[38,24] := -1.32375109;
      FC_W[38,25] := 0.04513154;
      FC_W[38,26] := 1.67587698;
      FC_W[38,27] := -0.60315883;
      FC_W[38,28] := 0.26211092;
      FC_W[38,29] := 0.19600734;
      FC_W[38,30] := 0.12759703;
      FC_W[38,31] := -0.80153352;
      FC_W[39,0] := -0.26302251;
      FC_W[39,1] := -0.13630611;
      FC_W[39,2] := -0.42582512;
      FC_W[39,3] := 1.35046661;
      FC_W[39,4] := 0.01697250;
      FC_W[39,5] := 0.46786672;
      FC_W[39,6] := 0.49501494;
      FC_W[39,7] := 0.76843983;
      FC_W[39,8] := 0.11361471;
      FC_W[39,9] := -0.69949502;
      FC_W[39,10] := 2.98522973;
      FC_W[39,11] := -0.60766679;
      FC_W[39,12] := 0.50049680;
      FC_W[39,13] := 0.03772873;
      FC_W[39,14] := 1.23203897;
      FC_W[39,15] := -0.50727296;
      FC_W[39,16] := -0.01674953;
      FC_W[39,17] := 0.65698963;
      FC_W[39,18] := -1.38105071;
      FC_W[39,19] := -1.02741539;
      FC_W[39,20] := -0.30104086;
      FC_W[39,21] := -0.84942061;
      FC_W[39,22] := -2.26705384;
      FC_W[39,23] := 0.34730250;
      FC_W[39,24] := 0.08819789;
      FC_W[39,25] := -0.56604064;
      FC_W[39,26] := 0.36780006;
      FC_W[39,27] := 0.00000264;
      FC_W[39,28] := -0.93792969;
      FC_W[39,29] := 0.56323957;
      FC_W[39,30] := 0.57272154;
      FC_W[39,31] := 0.84531051;
      FC_B[0] := 0.22904585;
      FC_B[1] := -0.32124424;
      FC_B[2] := -0.41430396;
      FC_B[3] := 0.23817410;
      FC_B[4] := 0.44676143;
      FC_B[5] := 0.05166011;
      FC_B[6] := -0.24827445;
      FC_B[7] := 0.02050643;
      FC_B[8] := -0.16593719;
      FC_B[9] := -0.19699521;
      FC_B[10] := -0.51350182;
      FC_B[11] := 0.38616806;
      FC_B[12] := -0.58952403;
      FC_B[13] := -0.46169797;
      FC_B[14] := 0.10238413;
      FC_B[15] := -0.37535465;
      FC_B[16] := 0.00366738;
      FC_B[17] := -0.21541971;
      FC_B[18] := 0.67242295;
      FC_B[19] := -1.18966842;
      FC_B[20] := -0.31347767;
      FC_B[21] := 0.14605546;
      FC_B[22] := -0.99858981;
      FC_B[23] := -0.68530029;
      FC_B[24] := -0.54384995;
      FC_B[25] := -0.55743998;
      FC_B[26] := -1.40273142;
      FC_B[27] := 0.84184837;
      FC_B[28] := 0.03169463;
      FC_B[29] := 1.14109719;
      FC_B[30] := -1.00650537;
      FC_B[31] := -1.22086596;
      FC_B[32] := -0.98691547;
      FC_B[33] := -1.37902105;
      FC_B[34] := -1.34311986;
      FC_B[35] := -0.70222050;
      FC_B[36] := 0.03677494;
      FC_B[37] := -0.62728751;
      FC_B[38] := 0.11721312;
      FC_B[39] := 0.56657410;

END_DATA_BLOCK
